Fanuc KAREL source: KF00078.KL

PROGRAM KF00078
%NOLOCKGROUP
%ENVIRONMENT STRNG
VAR
  I: INTEGER
  J: INTEGER
  X: REAL
  Y: REAL
  B: BOOLEAN
  C: BOOLEAN
  TXT: STRING[80]
  TXT2: STRING[80]
  AI: ARRAY[4] OF INTEGER
  BI: ARRAY[4] OF INTEGER
  P: XYZWPR
  JP: JOINTPOS
  PF: POSITION
  V1: VECTOR
  V2: VECTOR
  STATUS: INTEGER
BEGIN
  TXT = '12'
  TXT2 = '2'
  I = 12
  X = 2.5
  CNV_REAL_STR(X, 8, 2, TXT)
END KF00078
